// TIA Portal V20 export
Screen "principal"  800x420, Number=2
  ScreenLayer 
    IOField "I/O field_1" at 327,20 size 111x73  DataFormat=Decimal, FormatPattern=9999, Mode=InOutput
      ProcessValue := CONT1
    Button "Button_1" at 116,49 size 96x32  Mode=Text, TextOff="Marxa", TextOn="Text"
      on Press: SetBitWhileKeyPressed(Tag := Marxa, Bit := 0)
    Button "Button_2" at 113,104 size 96x32  Mode=Text, TextOff="Paro", TextOn="Text"
      on Press: SetBitWhileKeyPressed(Tag := Paro, Bit := 0)
    Button "Button_3" at 541,37 size 96x32  Mode=Text, TextOff="Reset", TextOn="Text"
      on Press: SetTag(Tag := CONT1, Value := 0)
    TextField "Text field_1" at 348,239 size 26x20  Text="M1"
    Group "Group_1"
      SymbolLibrary "Symbol library_1" at 304,104 size 120x120  Rotation=Angle0
      Group "Group"
        Circle "Circle_2" at 335,142 size 38x38
          RangeAppearanceAnimation "RangeAppearanceAnimation"
            tag KM1
            0..0: back #ff0000, fore #181c31
            1..1: back #00ff00, fore #181c31
        Circle "Circle_1" at 335,142 size 38x38
          RangeAppearanceAnimation "RangeAppearanceAnimation"
            tag alarma
            0..0: back #808080, fore #181c31
            1..1: back #ff0000, fore #181c31, flashing
          SingleBitVisibilityAnimation "VisibilityAnimation"
            tag alarma
